(* IEC 61131-3 sources: CS_4_Aufzugsteuerung/src/Stations/CP112/Steuerung/Class/BusInterfaceVARAN (part 2) *)

END_FUNCTION

FUNCTION VIRTUAL GLOBAL BusInterfaceVARAN::UpdateDO
	VAR_INPUT
		pCmd 	            : ^CmdStruct;
		presult 	        : ^results;
	END_VAR
  VAR
    pUPDATEDOCfg      : ^t_UpdateDOCfg;
    pCurrentDO        : ^t_DOCfg;
    changed           : BOOL;

    p_DOSettingsRd    : ^t_VaranDOSettingsRd;
    p_DOSettingsWr    : ^t_VaranDOSettingsWr;
    p_DOSettingsRdWr  : ^t_VaranDOSettingsRdWr;
  END_VAR

  changed := false;
  pUPDATEDOCfg := ((pCmd^.aPara[0])$^t_UpdateDOCfg);

  pResult^.uiLng := 4;

  if CheckHandle(Handle:= pUPDATEDOCfg^.Handle) then

    pCurrentDO := (pUPDATEDOCfg^.Handle)$^t_DOCfg;

    // Check if parameters were changed
    // Read Object
    if pCurrentDO^.RDWR = _BUS_IF_READ then

      if pCurrentDO^.lengthRead <> pUPDATEDOCfg^.ud_length_read  then
        // Check that new DO length is smaller then max DO length
        if pCurrentDO^.maxLengthRead >= pUPDATEDOCfg^.ud_length_read  then
          pCurrentDO^.lengthRead := pUPDATEDOCfg^.ud_length_read;
          changed := true;
        else
          pResult^.aData[0]$t_BusIFRetvalErrorcode := _BUS_IF_RETVAL_ERROR_UPDATEDO_DOLENGTH;
          return;
        end_if;
      end_if;

      if pCurrentDO^.AddrOffsetRead <>  pUPDATEDOCfg^.ud_addressoff_read then
        pCurrentDO^.AddrOffsetRead := pUPDATEDOCfg^.ud_addressoff_read;
        changed := true;
      end_if;

    // Write Object
    elsif pCurrentDO^.RDWR = _BUS_IF_WRITE then

      if pCurrentDO^.lengthWrite <> pUPDATEDOCfg^.ud_length_write  then
        // Check that new DO length is smaller then max DO length
        if pCurrentDO^.maxLengthWrite >= pUPDATEDOCfg^.ud_length_write  then
          pCurrentDO^.lengthWrite := pUPDATEDOCfg^.ud_length_write;
          changed := true;
        else
          pResult^.aData[0]$t_BusIFRetvalErrorcode := _BUS_IF_RETVAL_ERROR_UPDATEDO_DOLENGTH;
          return;
        end_if;
      end_if;

      if pCurrentDO^.AddrOffsetWrite <>  pUPDATEDOCfg^.ud_addressoff_write then
        pCurrentDO^.AddrOffsetWrite := pUPDATEDOCfg^.ud_addressoff_write;
        changed := true;
      end_if;

    // Read Write Object
    else

      if pCurrentDO^.lengthRead <> pUPDATEDOCfg^.ud_length_read  then
        // Check that new DO length is smaller then max DO length
        if pCurrentDO^.maxLengthRead >= pUPDATEDOCfg^.ud_length_read  then
          pCurrentDO^.lengthRead := pUPDATEDOCfg^.ud_length_read;
          changed := true;
        else
          pResult^.aData[0]$t_BusIFRetvalErrorcode := _BUS_IF_RETVAL_ERROR_UPDATEDO_DOLENGTH;
          return;
        end_if;
      end_if;

      if pCurrentDO^.AddrOffsetRead <>  pUPDATEDOCfg^.ud_addressoff_read then
        pCurrentDO^.AddrOffsetRead := pUPDATEDOCfg^.ud_addressoff_read;
        changed := true;
      end_if;

      if pCurrentDO^.lengthWrite <> pUPDATEDOCfg^.ud_length_write  then
        // Check that new DO length is smaller then max DO length
        if pCurrentDO^.maxLengthWrite >= pUPDATEDOCfg^.ud_length_write  then
          pCurrentDO^.lengthWrite := pUPDATEDOCfg^.ud_length_write;
          changed := true;
        else
          pResult^.aData[0]$t_BusIFRetvalErrorcode := _BUS_IF_RETVAL_ERROR_UPDATEDO_DOLENGTH;
          return;
        end_if;
      end_if;

      if pCurrentDO^.AddrOffsetWrite <>  pUPDATEDOCfg^.ud_addressoff_write then
        pCurrentDO^.AddrOffsetWrite := pUPDATEDOCfg^.ud_addressoff_write;
        changed := true;
      end_if;

    end_if;

    if b_PayloadSupport then
      if changed then
        // Update Address and length
        // Read Object
        if pCurrentDO^.RDWR = _BUS_IF_READ then

          ChangeDOLengthOffset( ud_DOHandle     := pCurrentDO^.pHandle$UDINT
                              , ud_offset_read  := pCurrentDO^.AddrOffsetRead
                              , ud_length_read  := pCurrentDO^.lengthRead);

        // Write Object
        elsif pCurrentDO^.RDWR = _BUS_IF_WRITE then

          ChangeDOLengthOffset( ud_DOHandle     := pCurrentDO^.pHandle$UDINT
                              , ud_offset_write := pCurrentDO^.AddrOffsetWrite
                              , ud_length_write := pCurrentDO^.lengthWrite);

        // Read Write Object
        else
          ChangeDOLengthOffset( ud_DOHandle     := pCurrentDO^.pHandle$UDINT
                              , ud_offset_read  := pCurrentDO^.AddrOffsetRead
                              , ud_length_read  := pCurrentDO^.lengthRead
                              , ud_offset_write := pCurrentDO^.AddrOffsetWrite
                              , ud_length_write := pCurrentDO^.lengthWrite);
        end_if;
      end_if;
    elsif pCurrentDO^.IsLongDO = FALSE then

      // Update Address and length and Reset DO
      // Read Object
      if pCurrentDO^.RDWR = _BUS_IF_READ then

        p_DOSettingsRd    := pCurrentDO^.pDataRead$^t_VaranDOSettingsRd  - VM_DO_OFFSET_RD;

        p_DOSettingsRd^.ud_Address                := DeviceAddress + pCurrentDO^.AddrOffsetRead;
        p_DOSettingsRd^.us_ByteCnt                := pCurrentDO^.lengthRead$USINT;
        pCurrentDO^.pHandle^.usLengthofExpAnswer  := sizeof(t_VaranDOSettingsRd.us_Command) + pCurrentDO^.lengthRead;

        ResetDataObject(p_handleDO:=  pCurrentDO^.pHandle
                      , us_state  :=  pCurrentDO^.pHandle^.ucCtrlStat AND 3         // don't change run status, just recalculate the retry timeout here
                      , ud_bytes  :=  pCurrentDO^.lengthRead);

      // Write Object
      elsif pCurrentDO^.RDWR = _BUS_IF_WRITE then

        p_DOSettingsWr    := pCurrentDO^.pDataWrite$^t_VaranDOSettingsWr - VM_DO_OFFSET_WR;

        p_DOSettingsWr^.ud_Address              := DeviceAddress + pCurrentDO^.AddrOffsetWrite;
        p_DOSettingsWr^.us_ByteCnt              := pCurrentDO^.lengthWrite$USINT;
        pCurrentDO^.pHandle^.usSendBufferLength := sizeof(t_VaranDOSettingsWr) + pCurrentDO^.lengthWrite;

        ResetDataObject(p_handleDO:=  pCurrentDO^.pHandle
                      , us_state  :=  pCurrentDO^.pHandle^.ucCtrlStat AND 3         // don't change run status, just recalculate the retry timeout here
                      , ud_bytes  :=  pCurrentDO^.lengthWrite);

      // Read Write Object
      else
        p_DOSettingsRdWr  := pCurrentDO^.pDataWrite$^t_VaranDOSettingsRdWr - VM_DO_OFFSET_RDWR;

        p_DOSettingsRdWr^.ud_AddressRd := DeviceAddress + pCurrentDO^.AddrOffsetRead;
        p_DOSettingsRdWr^.ud_AddressWr := DeviceAddress + pCurrentDO^.AddrOffsetWrite;

        p_DOSettingsRdWr^.us_ByteCntRd  := pCurrentDO^.lengthRead$USINT;
        p_DOSettingsRdWr^.us_ByteCntWr  := pCurrentDO^.lengthWrite$USINT;

        pCurrentDO^.pHandle^.usLengthofExpAnswer  := sizeof(t_VaranDOSettingsRdWr.us_Command) + pCurrentDO^.lengthRead;
        pCurrentDO^.pHandle^.usSendBufferLength   := sizeof(t_VaranDOSettingsRdWr) + pCurrentDO^.lengthWrite;

        ResetDataObject(p_handleDO:=  pCurrentDO^.pHandle
                      , us_state  :=  pCurrentDO^.pHandle^.ucCtrlStat AND 3         // don't change run status, just recalculate the retry timeout here
                      , ud_bytes  :=  pCurrentDO^.lengthRead + pCurrentDO^.lengthWrite);

      end_if;
    else

      // change long DO

      // Update Address and length and Reset DO
      // Read Object
      if pCurrentDO^.RDWR = _BUS_IF_READ then

        pCurrentDO^.pLongDOSettings^.ud_Address      := DeviceAddress + pCurrentDO^.AddrOffsetRead;
        pCurrentDO^.pLongDOSettings^.ui_ByteCount0   := pCurrentDO^.lengthRead;
        pCurrentDO^.pLongDOSettings^.us_ByteCount1   := 0;
        pCurrentDO^.pHandle^.usSendBufferLength      := 16#FFFF;
        pCurrentDO^.pHandle^.usLengthofExpAnswer     := 16#FFFF;

      // Write Object
      elsif pCurrentDO^.RDWR = _BUS_IF_WRITE then

        pCurrentDO^.pLongDOSettings^.ud_Address      := DeviceAddress + pCurrentDO^.AddrOffsetWrite;
        pCurrentDO^.pLongDOSettings^.ui_ByteCount0   := pCurrentDO^.lengthWrite;
        pCurrentDO^.pLongDOSettings^.us_ByteCount1   := 0;
        pCurrentDO^.pHandle^.usSendBufferLength      := 16#FFFF;
        pCurrentDO^.pHandle^.usLengthofExpAnswer     := 16#FFFF;

      end_if;
    end_if;

    pResult^.aData[0]$t_BusIFRetvalErrorcode := _BUS_IF_RETVAL_OK;

  else
    pResult^.aData[0]$t_BusIFRetvalErrorcode := _BUS_IF_RETVAL_ERROR_INVALID_HANDLE;
  end_if;

END_FUNCTION

FUNCTION VIRTUAL GLOBAL BusInterfaceVARAN::UpdateMoveDO
	VAR_INPUT
		pCmd 	        : ^CmdStruct;
		presult 	    : ^results;
	END_VAR
  VAR
    pUPDATEDOCfg  : ^t_UpdateDOMoveCfg;
    pCurrentDO    : ^t_DOMoveCfg;
    sd_retval     : DINT;
  END_VAR

  pUPDATEDOCfg := ((pCmd^.aPara[0])$^t_UpdateDOMoveCfg);

  pResult^.uiLng := 4;

  if CheckMovHandle(Handle:= pUPDATEDOCfg^.Handle) then

    pCurrentDO := (pUPDATEDOCfg^.Handle)$^t_DOMoveCfg;

    // Check if length Parameter was passed
    // Length is used with Payload and without
    if (pUPDATEDOCfg^.ud_length_move <> 0) &
       pUPDATEDOCfg^.ud_length_move <> VM_DO_PROPERTY_INVALID  then
      // if the size is smaller than the maximum or if we don't have interrupted our own copy for the move command
      if (pUPDATEDOCfg^.ud_length_move <= pCurrentDO^.lengthMoveMax) | (us_SkippedWriteBlocks = 0) then
        pCurrentDO^.lengthMove := pUPDATEDOCfg^.ud_length_move;
      else
        pResult^.aData[0]$t_BusIFRetvalErrorcode := _BUS_IF_RETVAL_ERROR_UPDATEDO_DOLENGTH;
        return;
      end_if;
    end_if;

    if b_PayloadSupport then

      if  pUPDATEDOCfg^.ud_handle_source <> 0 &
          pUPDATEDOCfg^.ud_handle_source <> VM_DO_PROPERTY_INVALID  then

        pCurrentDO^.sourceDOHandle := pUPDATEDOCfg^.ud_handle_source;
      end_if;

      if  pUPDATEDOCfg^.ud_addressoff_source <> VM_DO_PROPERTY_INVALID  then  // 0 is valid offset

        pCurrentDO^.sourceDOOffset := pUPDATEDOCfg^.ud_addressoff_source;
      end_if;

      if  pUPDATEDOCfg^.ud_handle_dest <> 0 &
          pUPDATEDOCfg^.ud_handle_dest <> VM_DO_PROPERTY_INVALID  then

        pCurrentDO^.destDOHandle := pUPDATEDOCfg^.ud_handle_dest;
      end_if;

      if  pUPDATEDOCfg^.ud_addressoff_dest <> VM_DO_PROPERTY_INVALID  then  // 0 is valid offset

        pCurrentDO^.destDOOffset := pUPDATEDOCfg^.ud_addressoff_dest;
      end_if;

      sd_retval := ChangeMovDOLengthOffset( ud_MovDOHandle              := pCurrentDO^.pHandle$UDINT
                                          , ud_SourceReadDOHandle       := pCurrentDO^.sourceDOHandle
                                          , ud_SourceReadOffset         := pCurrentDO^.sourceDOOffset
                                          , ud_DestinationWriteDOHandle := pCurrentDO^.destDOHandle
                                          , ud_DestinationWriteOffset   := pCurrentDO^.destDOOffset
                                          , ud_LengthMove               := pCurrentDO^.lengthMove);

      if sd_retval then
        pResult^.aData[0]$t_BusIFRetvalErrorcode := _BUS_IF_RETVAL_ERROR_UPDATE_MOVE_DO_FAILED;
      else
        pResult^.aData[0]$t_BusIFRetvalErrorcode := _BUS_IF_RETVAL_OK;
      end_if;

    else

      if pUPDATEDOCfg^.p_sourcedata <> nil &
         pUPDATEDOCfg^.p_sourcedata <> VM_DO_PROPERTY_INVALID then

        pCurrentDO^.pSourceDOData := pUPDATEDOCfg^.p_sourcedata;
      end_if;

      if pUPDATEDOCfg^.p_destdata   <> nil &
         pUPDATEDOCfg^.p_destdata   <> VM_DO_PROPERTY_INVALID then

        pCurrentDO^.pDestDOData := pUPDATEDOCfg^.p_destdata;
      end_if;

      pCurrentDO^.p_MovSettings^.ud_AddressSrc  := pCurrentDO^.pSourceDOData$UDINT;
      pCurrentDO^.p_MovSettings^.ud_AddressDest := pCurrentDO^.pDestDOData$UDINT;
      pCurrentDO^.p_MovSettings^.ui_ByteCnt     := pCurrentDO^.lengthMove;

      pResult^.aData[0]$t_BusIFRetvalErrorcode := _BUS_IF_RETVAL_OK;
    end_if;

  else
    pResult^.aData[0]$t_BusIFRetvalErrorcode := _BUS_IF_RETVAL_ERROR_INVALID_HANDLE;
  end_if;

END_FUNCTION

FUNCTION VIRTUAL GLOBAL BusInterfaceVARAN::SetDOPrescaler
	VAR_INPUT
		pCmd 	        : ^CmdStruct;
		presult 	    : ^results;
	END_VAR
  VAR
    pSetDOPreSCfg : ^t_SetDoPrescaler;
    pCurrentDO    : ^t_DOCfg;
  END_VAR

  pSetDOPreSCfg := ((pCmd^.aPara[0])$^t_SetDoPrescaler);

  pResult^.uiLng := 4;

  if CheckHandle(Handle:= pSetDOPreSCfg^.Handle) then

    pCurrentDO := (pSetDOPreSCfg^.Handle)$^t_DOCfg;

    if b_PayloadSupport then

      if SetPrescaler( ud_DOHandle   := pCurrentDO^.pHandle$UDINT
                     , Prescaler     := pSetDOPreSCfg^.Prescaler
                     , PrescalerCnt  := 0) = VARANMANAGER_OK then // Start at 0 = default We probably need to extend this functionality

        pResult^.aData[0]$t_BusIFRetvalErrorcode := _BUS_IF_RETVAL_OK;
      else
        pResult^.aData[0]$t_BusIFRetvalErrorcode := _BUS_IF_RETVAL_ERROR_INVALID_HANDLE;
      end_if;
    else

      pCurrentDO^.pHandle^.ucExePrescaler := pSetDOPreSCfg^.Prescaler;
      pCurrentDO^.PreScaler := pSetDOPreSCfg^.Prescaler;  // Saved as needed again as init value

      pResult^.aData[0]$t_BusIFRetvalErrorcode := _BUS_IF_RETVAL_OK;
    end_if;
  else

    pResult^.aData[0]$t_BusIFRetvalErrorcode := _BUS_IF_RETVAL_ERROR_INVALID_HANDLE;
  end_if;

END_FUNCTION

FUNCTION VIRTUAL GLOBAL BusInterfaceVARAN::SetTasksPrescaler
	VAR_INPUT
		pCmd 	            : ^CmdStruct;
		presult 	        : ^results;
	END_VAR
  VAR
  	pTaskPreScalerCfg : ^t_TaskPreScaler;
  END_VAR

  pTaskPreScalerCfg  := ((pCmd^.aPara[0])$^t_TaskPreScaler);

  pResult^.uiLng := 4;

  // Check passed data
  if pTaskPreScalerCfg^.Prescaler > 0 &
     pTaskPreScalerCfg^.Prescaler >= pTaskPreScalerCfg^.RtPreScanTrigger &
     pTaskPreScalerCfg^.Prescaler >= pTaskPreScalerCfg^.RtPostScanTrigger &
     pTaskPreScalerCfg^.Prescaler >= pTaskPreScalerCfg^.CyTrigger then

    TaskPrescaler.MaxCnt            := pTaskPreScalerCfg^.Prescaler;
    TaskPrescaler.RtPreScanTigger   := pTaskPreScalerCfg^.RtPreScanTrigger;
    TaskPrescaler.RtPostScanTrigger := pTaskPreScalerCfg^.RtPostScanTrigger;
    TaskPrescaler.CyTrigger         := pTaskPreScalerCfg^.CyTrigger;

    pResult^.aData[0]$t_BusIFRetvalErrorcode := _BUS_IF_RETVAL_OK;
  else
    pResult^.aData[0]$t_BusIFRetvalErrorcode := _BUS_IF_RETVAL_ERROR_INVALID_DATA;
  end_if;

END_FUNCTION

FUNCTION VIRTUAL GLOBAL BusInterfaceVARAN::ResetDO
	VAR_INPUT
		pCmd 	      : ^CmdStruct;
		presult 	  : ^results;
	END_VAR
  VAR
    pResetDOCfg : ^t_ResetDOCfg;
    pCurrentDO  : ^t_DOCfg;
  END_VAR

  pResult^.uiLng := 4;

  pResetDOCfg := ((pCmd^.aPara[0])$^t_ResetDOCfg);

  if CheckHandle(Handle:= pResetDOCfg^.Handle) then

    // Paylaod DO auto calculate Timeout when the DO changes
    // Just return OK
    if b_PayloadSupport = false then

      pCurrentDO := (pResetDOCfg^.Handle)$^t_DOCfg;

      // Reset DO
      // Read Object
      if (pCurrentDO^.RDWR = _BUS_IF_READ) then
        if pCurrentDO^.IsLongDO then
          ResetDataObject(p_handleDO :=  pCurrentDO^.pHandle
                          , us_state :=  VARAN_DO_NO_RUN         // No auto run, DO must be started by specific command
                          , ud_bytes :=  128);
        else
          ResetDataObject(p_handleDO :=  pCurrentDO^.pHandle
                          , us_state :=  VARAN_DO_NO_RUN         // No auto run, DO must be started by specific command
                          , ud_bytes :=  pCurrentDO^.lengthRead);
        end_if;

      // Write DO
      elsif pCurrentDO^.RDWR = _BUS_IF_WRITE then
        if pCurrentDO^.IsLongDO then
          ResetDataObject(p_handleDO :=  pCurrentDO^.pHandle
                          , us_state :=  VARAN_DO_NO_RUN         // No auto run, DO must be started by specific command
                          , ud_bytes :=  128);
        else
          ResetDataObject(p_handleDO :=  pCurrentDO^.pHandle
                          , us_state :=  VARAN_DO_NO_RUN         // No auto run, DO must be started by specific command
                          , ud_bytes :=  pCurrentDO^.lengthWrite);
        end_if;

      // Read Write DO
      else

        ResetDataObject(p_handleDO:=  pCurrentDO^.pHandle
                        , us_state  :=  VARAN_DO_NO_RUN         // No auto run, DO must be started by specific command
                        , ud_bytes  :=  pCurrentDO^.lengthRead + pCurrentDO^.lengthWrite);

      end_if;

    end_if;

    pResult^.aData[0]$t_BusIFRetvalErrorcode := _BUS_IF_RETVAL_OK;

  else
    pResult^.aData[0]$t_BusIFRetvalErrorcode := _BUS_IF_RETVAL_ERROR_INVALID_HANDLE;
  end_if;

END_FUNCTION

FUNCTION VIRTUAL GLOBAL BusInterfaceVARAN::AddTask
	VAR_INPUT
		pCmd 	        : ^CmdStruct;
		presult       : ^results;
	END_VAR
  VAR
  	pTASKCfg      : ^t_TaskCfg;
    _ud_dol_type  : UDINT;
  END_VAR

  presult^.uiLng    := 4;

  pTASKCfg := ((pCmd^.aPara[0])$^t_TaskCfg);

  // Check for null pointer
  if pTASKCfg^.pthis then

        // Convert passed t_BusIFPriority  to VARAN ud_dol_type
    if pTASKCfg^.Priority = _BUS_IF_ISO then
      _ud_dol_type := VARAN_DOL_ISO;
    else
      _ud_dol_type := VARAN_DOL_ASY;
    end_if;

    // Save the passed callback pointer according to the callOptions
    if pTASKCfg^.callOptions = CALL_OPTION_RT_PRESCAN then
      p_UserCalls.p_UpdateRt := (pTASKCfg^.pthis)$pVirtualBase;
    elsif pTASKCfg^.callOptions = CALL_OPTION_RT_POSTSCAN then
      p_UserCalls.p_UpDateRtPostScan := (pTASKCfg^.pthis)$pVirtualBase;
    elsif pTASKCfg^.callOptions = (CALL_OPTION_RT_PRESCAN or CALL_OPTION_RT_POSTSCAN) then
      p_UserCalls.p_UpdateRt := (pTASKCfg^.pthis)$pVirtualBase;
      p_UserCalls.p_UpDateRtPostScan := (pTASKCfg^.pthis)$pVirtualBase;
    else
      p_UserCalls.p_UpdateCy := (pTASKCfg^.pthis)$pVirtualBase;
    end_if;

    //Install Varantask
    VaranIn.AddVaranTask( _ud_dol_type,
                          p_this:=this,       // The callback pointer cannot be used directly because the class must be derived from VaranBase (p_VaranBase)
                          pTASKCfg^.callOptions);

    pResult^.aData[0]$t_BusIFRetvalErrorcode := _BUS_IF_RETVAL_OK;
  else
    pResult^.aData[0]$t_BusIFRetvalErrorcode := _BUS_IF_RETVAL_ERROR_INVALID_POINTER;
  end_if;

END_FUNCTION

FUNCTION VIRTUAL GLOBAL BusInterfaceVARAN::SetRunState
	VAR_INPUT
		pCmd 	            : ^CmdStruct;
		presult 	        : ^results;
	END_VAR
  VAR
  	pSETRUNSTATECfg   : ^t_SetRunStateCfg;
    pCurrentDO        : ^t_DOCfg;
    pCurrentDOMove    : ^t_DOMoveCfg;
    sd_RetVal         : DINT;
  END_VAR

  presult^.uiLng  := 4;

  pSETRUNSTATECfg := ((pCmd^.aPara[0])$^t_SetRunStateCfg);

  // Standard DO -----------------------------------------------------------------------------
  if CheckHandle(Handle:= pSETRUNSTATECfg^.Handle) then

    pCurrentDO := (pSETRUNSTATECfg^.Handle)$^t_DOCfg;

    if b_PayloadSupport then
      if pSETRUNSTATECfg^.NewRunState = _BUS_IF_RUN_STATE_SINGLE_RUN then
        pCurrentDO^.b_DOIsRunning.ContRun       := false; // Override cont run
        pCurrentDO^.b_DOIsRunning.StartRequest  := true;
        pResult^.aData[0]$t_BusIFRetvalErrorcode := _BUS_IF_RETVAL_OK;
      elsif pSETRUNSTATECfg^.NewRunState = _BUS_IF_RUN_STATE_CONT_RUN then
        if EnableDO(ud_DOHandle := pCurrentDO^.pHandle$UDINT) = VARANMANAGER_OK then

          //check if do must be added to list
          if bAddDOsToListSupport
          & pCurrentDO^.bsDoInsert.DOisInserted = FALSE
          & pCurrentDO^.bsDoInsert.RequestInsertLater = TRUE then
            sd_RetVal := MULTI_VARAN_IINSERTDOINTODOL(pCurrentDO^.pHandle$UDINT);
            pCurrentDO^.bsDoInsert.DOisInserted := TRUE;
          end_if;

          pResult^.aData[0]$t_BusIFRetvalErrorcode := _BUS_IF_RETVAL_OK;
        else
          pResult^.aData[0]$t_BusIFRetvalErrorcode := _BUS_IF_RETVAL_ERROR_INVALID_HANDLE;
        end_if;
        pCurrentDO^.b_DOIsRunning         := 0; // Override any singlerun states
        pCurrentDO^.b_DOIsRunning.ContRun := true;
      else
        if DisableDO(ud_DOHandle := pCurrentDO^.pHandle$UDINT) = VARANMANAGER_OK then
          pResult^.aData[0]$t_BusIFRetvalErrorcode := _BUS_IF_RETVAL_OK;
        else
          pResult^.aData[0]$t_BusIFRetvalErrorcode := _BUS_IF_RETVAL_ERROR_INVALID_HANDLE;
        end_if;
        pCurrentDO^.b_DOIsRunning         := 0;
      end_if;
    else
      if pSETRUNSTATECfg^.NewRunState = _BUS_IF_RUN_STATE_SINGLE_RUN then
        pCurrentDO^.pHandle^.ucCtrlStat := SetRunStatus(state:=VARAN_DO_SINGLE_RUN);
      elsif pSETRUNSTATECfg^.NewRunState = _BUS_IF_RUN_STATE_CONT_RUN then
        pCurrentDO^.pHandle^.ucCtrlStat := SetRunStatus(state:=VARAN_DO_CONT_RUN);
      else
        pCurrentDO^.pHandle^.ucCtrlStat := SetRunStatus(state:=VARAN_DO_NO_RUN);
      end_if;

      pResult^.aData[0]$t_BusIFRetvalErrorcode := _BUS_IF_RETVAL_OK;
    end_if;

  // Move DO ----------------------------------------------------------------------------------------
  elsif CheckMovHandle(Handle:= pSETRUNSTATECfg^.Handle) then

    pCurrentDOMove := (pSETRUNSTATECfg^.Handle)$^t_DOMoveCfg;

    if b_PayloadSupport then
      if pSETRUNSTATECfg^.NewRunState = _BUS_IF_RUN_STATE_SINGLE_RUN then
        pCurrentDOMove^.b_DOIsRunning.ContRun       := false; // Override cont run
        pCurrentDOMove^.b_DOIsRunning.StartRequest  := true;
        pResult^.aData[0]$t_BusIFRetvalErrorcode := _BUS_IF_RETVAL_OK;
      elsif pSETRUNSTATECfg^.NewRunState = _BUS_IF_RUN_STATE_CONT_RUN then
        if EnableDO(ud_DOHandle := pCurrentDOMove^.pHandle$UDINT) = VARANMANAGER_OK then
          pResult^.aData[0]$t_BusIFRetvalErrorcode := _BUS_IF_RETVAL_OK;
        else
          pResult^.aData[0]$t_BusIFRetvalErrorcode := _BUS_IF_RETVAL_ERROR_INVALID_HANDLE;
        end_if;
        pCurrentDOMove^.b_DOIsRunning         := 0; // Override any singlerun states
        pCurrentDOMove^.b_DOIsRunning.ContRun := true;
      else
        if DisableDO(ud_DOHandle := pCurrentDOMove^.pHandle$UDINT) = VARANMANAGER_OK then
          pResult^.aData[0]$t_BusIFRetvalErrorcode := _BUS_IF_RETVAL_OK;
        else
          pResult^.aData[0]$t_BusIFRetvalErrorcode := _BUS_IF_RETVAL_ERROR_INVALID_HANDLE;
        end_if;
        pCurrentDOMove^.b_DOIsRunning         := 0;
      end_if;
    else
      if pSETRUNSTATECfg^.NewRunState = _BUS_IF_RUN_STATE_SINGLE_RUN then
        pCurrentDOMove^.pHandle^.ucCtrlStat := SetRunStatus(state:=VARAN_DO_SINGLE_RUN);
      elsif pSETRUNSTATECfg^.NewRunState = _BUS_IF_RUN_STATE_CONT_RUN then
        pCurrentDOMove^.pHandle^.ucCtrlStat := SetRunStatus(state:=VARAN_DO_CONT_RUN);
      else
        pCurrentDOMove^.pHandle^.ucCtrlStat := SetRunStatus(state:=VARAN_DO_NO_RUN);
      end_if;

      pResult^.aData[0]$t_BusIFRetvalErrorcode := _BUS_IF_RETVAL_OK;
    end_if;

  else
    pResult^.aData[0]$t_BusIFRetvalErrorcode := _BUS_IF_RETVAL_ERROR_INVALID_HANDLE;
  end_if;

END_FUNCTION

FUNCTION VIRTUAL GLOBAL BusInterfaceVARAN::SetSyncData
	VAR_INPUT
		pCmd 	        : ^CmdStruct;
		presult 	    : ^results;
	END_VAR
  VAR
    pSYNCDATACfg  :  ^t_SyncData;
    i             : USINT;
  END_VAR

  presult^.uiLng  := 4;

  pSYNCDATACfg    := ((pCmd^.aPara[0])$^t_SyncData);

  i := pSYNCDATACfg^.us_sync_nr;

  if  i >= 0 &
      i <  4 then

    SyncData[i].us_sync_nr                := pSYNCDATACfg^.us_sync_nr;
    SyncData[i].sd_offset                 := pSYNCDATACfg^.sd_offset;
    SyncData[i].us_period_multiplier      := pSYNCDATACfg^.us_period_multiplier;
    SyncData[i].us_enable_frame_count     := pSYNCDATACfg^.us_enable_frame_count;
    SyncData[i].us_frame_count_threshold  := pSYNCDATACfg^.us_frame_count_threshold;
    SyncData[i].b_use_divider_sync        := pSYNCDATACfg^.b_use_divider_sync;

    bSetPll := TRUE;

    pResult^.aData[0]$t_BusIFRetvalErrorcode := _BUS_IF_RETVAL_OK;
  else
    pResult^.aData[0]$t_BusIFRetvalErrorcode := _BUS_IF_RETVAL_ERROR_INVALID_SYNC;
  end_if;

END_FUNCTION

FUNCTION VIRTUAL BusInterfaceVARAN::CheckHandle
	VAR_INPUT
		Handle 	    : UDINT;
	END_VAR
	VAR_OUTPUT
		IsOk 	      : BOOL;
	END_VAR
  VAR
    ListOffset  : UDINT;
  END_VAR

  IsOk := false;

  // Handle must be not nil and there must be elements in the array.
  if Handle & NrDO then
    ListOffset := (Handle - (#DOList[0])$UDINT);
    if ((ListOffset MOD sizeof(t_DOCfg)) = 0) & ((ListOffset/sizeof(t_DOCfg)) < NrDO) then
      IsOk := true;
    end_if;
  end_if;

END_FUNCTION

FUNCTION VIRTUAL BusInterfaceVARAN::CheckMovHandle
	VAR_INPUT
		Handle 	    : UDINT;
	END_VAR
	VAR_OUTPUT
		IsOk 	      : BOOL;
	END_VAR
  VAR
    ListOffset  : UDINT;
  END_VAR

  IsOk := false;

  // Handle must be not nil and there must be elements in the array.
  if Handle & NrDOMove then
    ListOffset := (Handle - (#DOListMove[0])$UDINT);
    if ((ListOffset MOD sizeof(t_DOMoveCfg)) = 0) & ((ListOffset/sizeof(t_DOMoveCfg)) < NrDOMove) then
      IsOk := true;
    end_if;
  end_if;

END_FUNCTION

FUNCTION VIRTUAL GLOBAL BusInterfaceVARAN::UpdateRetryCounter
  VAR
    i                 : USINT;
	  tempRetryCounter  : USINT;
    pDOElement        : ^t_DOCfg;
  END_VAR

  // Standard DOs --------------------------------------------------------------------------
  if NrDO then
    pDOElement := #DOList[0];
    for i := 0 to (NrDO - 1) do

      tempRetryCounter := GetRetryCounter(ud_DOHandle := pDOElement^.pHandle$UDINT);

      if ( tempRetryCounter <> pDOElement^.OldRetryCounter) then
        RetryCounter += TO_USINT( tempRetryCounter - pDOElement^.OldRetryCounter );
        pDOElement^.OldRetryCounter := tempRetryCounter;
      end_if;

      pDOElement += sizeof(t_DOCfg);
    end_for;
  end_if;

END_FUNCTION

FUNCTION BusInterfaceVARAN::BusInterfaceVARAN
	VAR_OUTPUT
		ret_code 	: ConfStates;
	END_VAR

  ui_PostInitIndex := 16#FFFF;

  // initialize with 0xff for invalid
  _memset(dest:=#SyncData, usByte:=16#FF, cntr:=sizeof(SyncData));

  if OS_CILGet(INTERFACE_VARANMANAGER, #pVaran) <> SYS_ERR_NONE then
    LogError("@0196 (BusInterfaceVARAN::BusInterfaceVARAN) Failed to get VARAN-CIL (interface to OS)!");
  end_if;

  b_LongDOsPossible := GetLongDOsPossible();

	ret_code := C_OK;

END_FUNCTION

FUNCTION VIRTUAL GLOBAL BusInterfaceVARAN::Varan_HwInterrupt
	VAR_INPUT
		ud_reason 	: UDINT;
		ud_data 	  : ^t_CallBackInterrupt;
	END_VAR
	VAR_OUTPUT
		sd_retval 	: DINT;
	END_VAR
  VAR
  	tempCmd     : CmdStruct;
    _result     : results;
  END_VAR;

  // Turn off DO's
  SetDOsOff();

  // Check for 0 pointer
  if p_UserCalls.p_Callback then
    // Call the corrosponding function in the operator class
    tempCmd.uiCmd := _BUS_IF_HWINTERRUPT;
    p_UserCalls.p_Callback^.pSvrChCmd.NewInst(#tempCmd,#_result);
  end_if;
  sd_retval := Varan_Base::Varan_HwInterrupt(ud_reason, ud_data);

END_FUNCTION

FUNCTION VIRTUAL BusInterfaceVARAN::LogErrorExt
	VAR_INPUT
		e_msg 	    : ^CHAR;
		p_extThis1 	: pVirtualBase;
		p_extThis2 	: pVirtualBase;
	END_VAR
  VAR
    sz_name     : ARRAY [ 0..255 ] OF CHAR;
    MyMsg       : ARRAY [0..599] OF CHAR;
  END_VAR

  if p_extThis1 = nil then
    p_extThis1 := this;
  end_if;

  if p_extThis2 then
    _GetObjName( p_extThis2, #sz_name[ 0 ] );
#ifdef HWC_LimitObjName
    HWC_LimitObjName(#sz_name[ 0 ]);
#endif
    _strncpy(dest:=#MyMsg[0], src:=e_msg, max:=200);
    _strcat( dest:=#MyMsg[0], src:=" ");
    _strcat( dest:=#MyMsg[0], src:=#sz_name[0]);

#ifdef HWC_LogError
    HWC_LogError(p_extThis1, #MyMsg[0]);
#endif

  else
#ifdef HWC_LogError
    HWC_LogError(p_extThis1, e_msg);
#endif
  end_if;

END_FUNCTION

FUNCTION VIRTUAL BusInterfaceVARAN::InstallCallbackObject
	VAR_OUTPUT
		sd_retval 	: DINT;
	END_VAR

  // we don't install the callback here (1st init). it's installed in the 2nd init, because in the first init the operator may set us to required
  sd_retval := VARANMANAGER_OK;

END_FUNCTION

FUNCTION VIRTUAL BusInterfaceVARAN::GetLongDOsPossible
	VAR_OUTPUT
		LongDOsPossible 	  : BOOL;
	END_VAR
  VAR
    pSPCIInfo           : ^LSL_SPCIINFO;
  	p_sigmatek_devinfo 	: ^PCICONFDATA;
    p_NodeInfo          : ^LSL_VARANNODEINFO;
    ManagerNodeString   : USINT;
    ud_VMNodeHandle     : UDINT;
    s_NodeInfo          : LSL_VARANNODEINFO;
    sd_retval           : DINT;
  END_VAR

  LongDOsPossible := FALSE;

  // check if long DOs are supported by VARAN Manager. Version of wb_varan_manager_control_status_info (Device Type x"0212" of info block) has to be >= 16#25.
  if OS_CILGET( "PCICONFIG", #pSPCIInfo ) =  SYS_ERR_NONE then
    p_sigmatek_devinfo 	:= SPCIINFO_FINDDEVICE(0x0212, 0);
    if p_sigmatek_devinfo = NIL then
      p_sigmatek_devinfo 	:= SPCIINFO_FINDDEVICE(0x0214, 0); //check for new varan interface
    end_if;
    // check if the Manager supports LongDOs
    if p_sigmatek_devinfo & (p_sigmatek_devinfo^.Version >= 16#25) then
      LongDOsPossible := TRUE;
    else
      // we don't get the device at a c-ipc, because it's a pci plug-in card
      if pVaran & (_WhoAmI = DESTPLC_C_IPC) then
        // now check the platform and the corresponding fpga version

        //get manager node info from os
        ManagerNodeString := 0;

        //call OS - function (must be OS-funciton because of error handling)
        if b_PayloadSupport then
          // Get the Handle of the VM
          sd_retval := MULTI_VARAN_iGetNodeHandle(udManagerNumber := ud_VaranManagerNr
                                                , pszHardwarePath := #ManagerNodeString
                                                , phNodeHandle    := #ud_VMNodeHandle);

          if sd_retval = VARANMANAGER_OK then
            p_NodeInfo := #s_NodeInfo;
            sd_retval := MULTI_VARAN_iGetNodeInformation( hNodeHandle := ud_VMNodeHandle
                                                        , psNodeInfo  := p_NodeInfo);     // Pass a pointer to the buffer into which the data will be written, instead of getting a pointer to te data
          end_if;

        else
          sd_retval := VARAN_iGetNodeInfo(uiManager	:= ud_VaranManagerNr
                                        , pucNode	  := #ManagerNodeString
                                        , pNodeInfo	:= #p_NodeInfo
                                        );
        end_if;

        if	( sd_retval = VARANMANAGER_OK ) & p_NodeInfo then
          case p_NodeInfo^.uiDeviceID of
            1000: // VM051    >= 1.6
              if p_NodeInfo^.ucFPGAVersion >= 16#16 then
                LongDOsPossible := TRUE;
              end_if;

            1030, // VM052    >= 1.4
            1150: // VM052-1  same fpga file
              if p_NodeInfo^.ucFPGAVersion >= 16#14 then
                LongDOsPossible := TRUE;
              end_if;

            1031: // VM052H   not necessary, this card doesn't work on a C-IPC (created for customer specific hardware)

            1044: // VMC052   >= 1.3
              if p_NodeInfo^.ucFPGAVersion >= 16#13 then
                LongDOsPossible := TRUE;
              end_if;

            1063, // VM052-3  >= 1.4
            1093: // VM053    same fpga file
              if p_NodeInfo^.ucFPGAVersion >= 16#14 then
                LongDOsPossible := TRUE;
              end_if;

            1080: // VM052-4  no fpga available

          end_case;
        end_if;
      end_if;
    end_if;
  end_if;

END_FUNCTION

FUNCTION VIRTUAL GLOBAL BusInterfaceVARAN::Varan_HwSubBusReady
	VAR_INPUT
		ud_data 	  : UDINT;
	END_VAR
	VAR_OUTPUT
		sd_retval 	: DINT;
	END_VAR
  VAR
  	tempCmd     : CmdStruct;
    _result     : results;
  END_VAR

  // Check for 0 pointer
  if p_UserCalls.p_Callback then
    // Call the corresponding function in the operator class
    tempCmd.uiCmd := _BUS_IF_HWSUB_BUS_READY;
    p_UserCalls.p_Callback^.pSvrChCmd.NewInst(#tempCmd,#_result);

    sd_retval := _result.aData[0]$DINT;
  else
    sd_retval := 0;
  end_if;

END_FUNCTION

FUNCTION VIRTUAL GLOBAL BusInterfaceVARAN::State::NewInst
	VAR_INPUT
		pPara 	    : ^CmdStruct;
		pResult 	  : ^Results;
	END_VAR
	VAR_OUTPUT
		ret_code 	  : IprStates;
	END_VAR
  VAR
  	tempCmd     : CmdStruct;
    _result     : results;
    // local variables for the Requested HWTString
    pStr_HWTRequested       : ^CHAR;
    us_HWTRequestedCurrIndex: USINT;
    pStr_HWTreenEntry       : ^CHAR;
    ud_HWCRetcode           : t_HWCRetvalReturnCode;
    b_CallThisModule        : BOOL;
  END_VAR

  pStr_HWTRequested         := NIL;
  us_HWTRequestedCurrIndex  := 0;
  pStr_HWTreenEntry         := NIL;
  ud_HWCRetcode             := _HWC_RETVAL_ERROR;
  b_CallThisModule          := TRUE;

	ret_code := READY;

  CASE pPara^.uiCmd OF
//**********************************************************************************************************************************************************
    CMD_POST_INIT_RT_READY:
      // check if operator is ready
      tempCmd.uiCmd := _BUS_IF_POST_INIT_RT_READY;
      ret_code := p_UserCalls.p_Callback^.pSvrChCmd.NewInst(#tempCmd, #_result);

      if bSimulateSDIASManager then

        // if we got an error => return it
        if eSdiasManagerInitSSW = _ErrorOccured then
          ret_code := ERROR;

        //if we're not ready, return busy
        elsif eSdiasManagerInitSSW <> _InitFinished then
          ret_code := BUSY;
        end_if;

      end_if;

//**********************************************************************************************************************************************************
    CMD_GET_HARDWARE_DIAGNOSIS:

      pResult^.aData$t_HWCGetHardwareDiagnosisOut.retcode := _HWC_RETVAL_ERROR_CLASS_NOT_ONLINE;
      ret_code := ERROR;

      pResult^.aData[0]$t_HWCGetHardwareDiagnosisOut.retcode := _HWC_RETVAL_ERROR;

      pStr_HWTRequested := pPara^.aPara[0]$t_HWCGetHardwareDiagnosisIn.pStr_HardewareTreeEntry;

      // Check HWT String
      if pStr_HWTRequested then

        us_HWTRequestedCurrIndex  := pPara^.aPara[0]$t_HWCGetHardwareDiagnosisIn.us_current_index;

        // Check for any Escape sequence
        if (pStr_HWTRequested + us_HWTRequestedCurrIndex)^ and HWT_ESCAPE_SEQU then

          // Check if current index + 1 is valid, pStr_HWTRequested^ + 1 for extra byte of length
          if (us_HWTRequestedCurrIndex + 1) <= (pStr_HWTRequested$^UINT^ + 1) then
            // Update Current index to next position = Place of SDIAS Module
            pPara^.aPara[0]$t_HWCGetHardwareDiagnosisIn.us_current_index   += 1;
            pPara^.aPara[0]$t_HWCGetHardwareDiagnosisIn.us_current_length  -= 1;

            if p_UserCalls.p_Callback then
              ret_code := p_UserCalls.p_Callback^.pSvrChCmd.NewInst(pPara,pResult); //Pass on command to connected extension module
            end_if;

          end_if;

        else
          ret_code := Varan_Base::State.NewInst(pPara, pResult);  // Pass on command to base

          // Call conneceted Class for additional info
          if p_UserCalls.p_Callback then

            // Don't change retcode, may be not handled by extension modules.
            ud_HWCRetcode := pResult^.aData[0]$t_HWCGetHardwareDiagnosisOut.retcode;

            p_UserCalls.p_Callback^.pSvrChCmd.NewInst(pPara,pResult); //Pass on command to extension module

            pResult^.aData[0]$t_HWCGetHardwareDiagnosisOut.retcode := ud_HWCRetcode;

          end_if;
        end_if;

      end_if;

//**********************************************************************************************************************************************************

    CMD_GET_HARDWARE_TREE_ENTRY:

      pResult^.aData$t_HWCGetHardwareTreeEntryOut.retcode := _HWC_RETVAL_ERROR_CLASS_NOT_ONLINE;
      ret_code            := ERROR;

      pStr_HWTRequested   := pPara^.aPara[0]$t_HWCGetHardwareTreeEntryIn.pStr_LastHardewareTreeEntry;

      b_CallThisModule    := TRUE;

      // Check HWT String
      if pStr_HWTRequested & p_ObjectPath then

        // Compare string content
        if _memcmp( ptr1 := pStr_HWTRequested + 2,
                    ptr2 := p_ObjectPath +1,
                    cntr := p_ObjectPath^) = 0 then

          //Check if last call was to Base itself, Compare string length
          if (pStr_HWTRequested$^USINT^ = p_ObjectPath^) then

            //If last call was to base itself, don't call it this time
            b_CallThisModule := FALSE;

            // Last module called was the BusIF Object itself, next module is the 1st behind the extension module
            pPara^.aPara[0]$t_HWCGetHardwareTreeEntryIn.pStr_LastHardewareTreeEntry := NIL;

            if p_UserCalls.p_Callback then
              ret_code := p_UserCalls.p_Callback^.pSvrChCmd.NewInst(pPara,pResult); //Pass on command to extension module

              // if we should quit treating this module special => use standard behavior
              if ret_code = QUIT then
                ret_code := Varan_Base::State.NewInst(pPara,pResult); //Pass on command to base
              end_if;

            else
              pResult^.aData[0]$t_HWCGetHardwareTreeEntryOut.retcode := _HWC_RETVAL_OK_END_OF_LIST;
            end_if;

          elsif (pStr_HWTRequested$^USINT^ > p_ObjectPath^ + 1) then // Must be at least 2 Byte larger, ESCAPE Sequence + Place

            // Check escape sequence
            if ( (pStr_HWTRequested + (p_ObjectPath^) + 2 )^ AND HWT_ESCAPE_SEQU) then // First place after extension module Itself is escape sequence + 1 for addional length byte
              // Last Module must have been a Module behind an extension module

              //If last call was to base itself, don't call it this time
              b_CallThisModule := FALSE;

              // Update index
              pPara^.aPara[0]$t_HWCGetHardwareTreeEntryIn.us_current_index  := p_ObjectPath^ + 3; // Second place after BUSIF Itself is place + 1 for addional length byte
              pPara^.aPara[0]$t_HWCGetHardwareTreeEntryIn.us_current_length := pStr_HWTRequested^ - p_ObjectPath^ - 1;

              //If we have a extension module
              if p_UserCalls.p_Callback then
                ret_code := p_UserCalls.p_Callback^.pSvrChCmd.NewInst(pPara,pResult); //Pass on command to extension module
              else
                ret_code := READY;
                pResult^.aData[0]$t_HWCGetHardwareTreeEntryOut.retcode := _HWC_RETVAL_OK_END_OF_LIST;
              end_if;
            end_if;
          end_if;
        end_if;
      end_if;

      if b_CallThisModule then

        ret_code := Varan_Base::State.NewInst(pPara, pResult);  // Pass on command to base

        // Call conneceted Class for additional info
        if p_UserCalls.p_Callback &
           pResult^.aData[0]$t_HWCGetHardwareTreeEntryOut.pStr_NextHardewareTreeEntry then

          // Update with Requested HWT String with the one returned from Varanbase
          pPara^.aPara[0]$t_HWCGetHardwareTreeEntryIn.pStr_LastHardewareTreeEntry := pResult^.aData[0]$t_HWCGetHardwareTreeEntryOut.pStr_NextHardewareTreeEntry;

          // Don't change retcode, may be not handled by extension modules.
          ud_HWCRetcode := pResult^.aData[0]$t_HWCGetHardwareTreeEntryOut.retcode;

          p_UserCalls.p_Callback^.pSvrChCmd.NewInst(pPara,pResult); //Pass on command to extension module

          pResult^.aData[0]$t_HWCGetHardwareTreeEntryOut.retcode := ud_HWCRetcode;
        end_if;
      end_if;

//**********************************************************************************************************************************************************

   CMD_GET_HW_TIMESTAMP:
      // forward to VM
      ret_code := VaranIn.NewInst(pPara, pResult);

//**********************************************************************************************************************************************************

   CMD_HWC_REQ_PLLNS_REGULATION:
      // forward to VM
      ret_code := VaranIn.NewInst(pPara, pResult);

//**********************************************************************************************************************************************************

  ELSE
    // unknown commands are forwarded to the base
    ret_code := Varan_Base::State.NewInst(pPara, pResult);
  END_CASE;

END_FUNCTION

FUNCTION VIRTUAL GLOBAL BusInterfaceVARAN::GetDeviceID
	VAR_OUTPUT
		output 	: UDINT;
	END_VAR

  output := DeviceIDDiagnosis;

END_FUNCTION

FUNCTION VIRTUAL GLOBAL BusInterfaceVARAN::GetPayloadSupportState
	VAR_OUTPUT
		dRetCode 	: DINT;
	END_VAR

  dRetCode := b_PayloadSupport;

END_FUNCTION

FUNCTION VIRTUAL BusInterfaceVARAN::AddSDORequest
	VAR_INPUT
		pCmdSvr 	: ^SvrChCmd;
		Command 	: HINT;
		Offset 	: UDINT;
		Length 	: UDINT;
		pWriteBuf 	: ^void;
	END_VAR
	VAR_OUTPUT
		sd_retval 	: DINT;
	END_VAR

  // protect via mutex because this can be called from different task priorities
  OS_MT_WAIT(pv_MutexSDOs);

  // if the buffer is full, or the next element in the buffer is already in use
  if (SDOHandling.pWrite^.Command <> 0) then
    sd_retval := -2;
    OS_MT_SIGNAL(pv_MutexSDOs);
    return;
  end_if;

  if pCmdSvr = NIL then
    sd_retval := -3;
    return;
  end_if;

  if Length = 0 then
    sd_retval := -4;
  end_if;

  if Command =_BUS_IF_WRITE_VIA_SDO | Command = _BUS_IF_WRITE_VIA_SDO_CTRL then
    if pWriteBuf = NIL then
      sd_retval := -5;
      return;
    end_if;
  end_if;

  SDOHandling.pWrite^.pCallBackSvr  := pCmdSvr;
  SDOHandling.pWrite^.udLength      := Length;
  SDOHandling.pWrite^.udOffset      := Offset;
  SDOHandling.pWrite^.pWriteData    := pWriteBuf;
  // command is the last thing to store, because it indicates a complete entry
  SDOHandling.pWrite^.Command := Command;

  // we increment our used entries in the buffer (only for debugging)
  SDOHandling.EntriesUsed     += 1;

  // after we successfully added this SDO, set the write pointer to the next element
  if SDOHandling.pWrite = SDOHandling.pLastEntry then
    SDOHandling.pWrite := SDOHandling.pRingBufMemStart;
  else
    SDOHandling.pWrite += sizeof(t_SDORingBufEntry);
  end_if;

  sd_retval := 0;

  OS_MT_SIGNAL(pv_MutexSDOs);

END_FUNCTION

FUNCTION VIRTUAL BusInterfaceVARAN::CyclicSDOHandling
  VAR
		Length 	      : UDINT;
    pRingBufEntry : ^t_SDORingBufEntry;
    pCmdSvr       : ^SvrChCmd;
  	tempCmd       : CmdStruct;
    _result       : results;
    Offset : UDINT;
  END_VAR

  // protect via mutex because this can be called from different task priorities
  OS_MT_WAIT(pv_MutexSDOs);

  //If there is some work todo
  if SDOHandling.EntriesUsed then

    if SDOHandling.pActEntry & SDOHandling.pActEntry^.Command <> 0 then

      pRingBufEntry := SDOHandling.pActEntry;

      //State = 0 ... Start SDO access, 1 ... Get SDO access data and stop SDO
      if SDOHandling.pActEntry^.udState = 0 then

        Length := SDOHandling.pActEntry^.udLength;
        Offset := SDOHandling.pActEntry^.udOffset;

        case SDOHandling.pActEntry^.Command of

          _BUS_IF_READ_VIA_SDO:

            if ChangeAsyRd(Offset:=Offset$UINT,
                           Length:=Length$USINT,
                           RunState:=_BUS_IF_RUN_STATE_CONT_RUN,
                           bIsCtrlACC := FALSE) = FALSE then
              LogError("@009B (BusInterfaceVARAN::CyclicSDOHandling) Error occured at starting the MEM ReadDO");
            end_if;

            SDOHandling.pActEntry^.udState := 1;

          _BUS_IF_READ_VIA_SDO_CTRL:

            if ChangeAsyRd(Offset:=Offset$UINT,
                           Length:=Length$USINT,
                           RunState:=_BUS_IF_RUN_STATE_CONT_RUN,
                           bIsCtrlACC := TRUE) = FALSE then
              LogError("@009B (BusInterfaceVARAN::CyclicSDOHandling) Error occured at starting the CTRL ReadDO");
            end_if;

            SDOHandling.pActEntry^.udState := 1;

          _BUS_IF_WRITE_VIA_SDO:

            _memcpy(ptr1:=AsyMemWriteDO.pData, ptr2:=SDOHandling.pActEntry^.pWriteData, cntr:=SDOHandling.pActEntry^.udLength);

            if ChangeAsyWr(Offset:=Offset$UINT,
                           Length:=Length$USINT,
                           RunState:=_BUS_IF_RUN_STATE_CONT_RUN,
                           bIsCtrlACC := FALSE) = FALSE then
              LogError("@009B (BusInterfaceVARAN::CyclicSDOHandling) Error occured at starting the MEM WriteDO");
            end_if;

            SDOHandling.pActEntry^.udState := 1;

          _BUS_IF_WRITE_VIA_SDO_CTRL:

            _memcpy(ptr1:=AsyCtrlWriteDO.pData, ptr2:=SDOHandling.pActEntry^.pWriteData, cntr:=SDOHandling.pActEntry^.udLength);

            if ChangeAsyWr(Offset:=Offset$UINT,
                           Length:=Length$USINT,
                           RunState:=_BUS_IF_RUN_STATE_CONT_RUN,
                           bIsCtrlACC := TRUE) = FALSE then
              LogError("@009B (BusInterfaceVARAN::CyclicSDOHandling) Error occured at starting the CTRL WriteDO");
            end_if;

            SDOHandling.pActEntry^.udState := 1;

        end_case;

      elsif SDOHandling.pActEntry^.udState = 1 then

        SDOHandling.EntriesUsed -= 1;

        // Call the corresponding function in the operator class
        tempCmd.uiCmd := _BUS_IF_SDO_RESPONSE;
        tempCmd.aPara[0] := SDOHandling.pActEntry^.Command$DINT;
        tempCmd.aPara[1] := SDOHandling.pActEntry^.udOffset$DINT;
        tempCmd.aPara[2] := SDOHandling.pActEntry^.udLength$DINT;

        tempCmd.aPara[3] := 0;

        case SDOHandling.pActEntry^.Command of

          _BUS_IF_READ_VIA_SDO:

            tempCmd.aPara[4] := AsyMemReadDO.pData$DINT;
            tempCmd.aPara[5] := AsyMemReadDO.Length;

          _BUS_IF_READ_VIA_SDO_CTRL:

            tempCmd.aPara[4] := AsyCtrlReadDO.pData$DINT;
            tempCmd.aPara[5] := AsyCtrlReadDO.Length;

          _BUS_IF_WRITE_VIA_SDO:

            tempCmd.aPara[4] := NIL$DINT;
            tempCmd.aPara[5] := 0;

          _BUS_IF_WRITE_VIA_SDO_CTRL:

            tempCmd.aPara[4] := NIL$DINT;
            tempCmd.aPara[5] := 0;

        end_case;

        pCmdSvr := pRingBufEntry^.pCallBackSvr;

        if pCmdSvr$pVirtualBase^.NewInst(#tempCmd, #_result) <> READY then
          LogError("@0099 (BusInterfaceVARAN::CyclicSDOHandling) SDO Error: Error of module at place 0x{0} while receiving the SDO reponse (which was an ErrorCode)");
        end_if;

        // the entry in the ringbuffer is free
        pRingBufEntry^.Command := 0;

        //Stop the DOs
        if ChangeAsyRd(Offset:=0,
                       Length:=0,
                       RunState:=_BUS_IF_RUN_STATE_NO_RUN,
                       bIsCtrlACC := TRUE) = FALSE then
          LogError("@0769 (BusInterfaceVARAN::CyclicSDOHandling) Error occured at starting the CTRL ReadDO");
        end_if;

        if ChangeAsyRd(Offset:=0,
                       Length:=0,
                       RunState:=_BUS_IF_RUN_STATE_NO_RUN,
                       bIsCtrlACC := FALSE) = FALSE then
          LogError("@076A (BusInterfaceVARAN::CyclicSDOHandling) Error occured at starting the MEM ReadDO");
        end_if;

        if ChangeAsyWr(Offset:=0,
                       Length:=0,
                       RunState:=_BUS_IF_RUN_STATE_NO_RUN,
                       bIsCtrlACC := TRUE) = FALSE then
          LogError("@076B (BusInterfaceVARAN::CyclicSDOHandling) Error occured at starting the CTRL WriteDO");
        end_if;

        if ChangeAsyWr(Offset:=0,
                       Length:=0,
                       RunState:=_BUS_IF_RUN_STATE_NO_RUN,
                       bIsCtrlACC := FALSE) = FALSE then
          LogError("@076D (BusInterfaceVARAN::CyclicSDOHandling) Error occured at starting the MEM WriteDO");
        end_if;

        SDOHandling.pActEntry^.udState := 0;

        // after we successfully added this SDO, set the read pointer to the next element
        if SDOHandling.pActEntry = SDOHandling.pLastEntry then
          SDOHandling.pActEntry := SDOHandling.pRingBufMemStart;
        else
          SDOHandling.pActEntry += sizeof(t_SDORingBufEntry);
        end_if;

      end_if;
    end_if;
  end_if;

  OS_MT_SIGNAL(pv_MutexSDOs);

END_FUNCTION

FUNCTION VIRTUAL BusInterfaceVARAN::ChangeAsyRd
	VAR_INPUT
		Offset 	: HINT;
		Length 	: USINT;
		RunState 	: t_BusIFRunState;
		bIsCtrlACC 	: BOOL;
	END_VAR
	VAR_OUTPUT
		Success 	: BOOL;
	END_VAR
  VAR
    dataUPDATEDO    : t_UpdateDOCfg;
  	tempCmd         : CmdStruct;
    _result         : results;
    dataSETRUNSTATE : t_SetRunStateCfg;
  END_VAR

  // if length = zero we may just want to stop the DO
  if Length then

    if bIsCtrlACC then
      AsyCtrlReadDO.Offset := Offset;
      AsyCtrlReadDO.Length := Length;

      dataUPDATEDO.Handle               := AsyCtrlReadDO.Handle;
      dataUPDATEDO.ud_addressoff_read   := AsyCtrlReadDO.Offset;
      dataUPDATEDO.ud_length_read       := AsyCtrlReadDO.Length;

    else
      AsyMemReadDO.Offset := Offset;
      AsyMemReadDO.Length := Length;

      dataUPDATEDO.Handle               := AsyMemReadDO.Handle;
      dataUPDATEDO.ud_addressoff_read   := AsyMemReadDO.Offset;
      dataUPDATEDO.ud_length_read       := AsyMemReadDO.Length;
    end_if;

    tempCmd.uiCmd         := _BUS_IF_UPDATE_DO;
    tempCmd.aPara[0]      := (#dataUPDATEDO)$DINT;

    CallCommand.NewInst(pPara:=#tempCmd, pResult:=#_result);
    if _result.aData[0]$t_BusIFRetvalErrorcode <> _BUS_IF_RETVAL_OK then
      LogError("@007C (BusInterfaceVARAN::ChangeAsyRd) Failed to change asynchron read access");
    end_if;
  end_if;

  // set runstate
  if bIsCtrlACC then
    dataSETRUNSTATE.Handle      := AsyCtrlReadDO.Handle;
  else
    dataSETRUNSTATE.Handle      := AsyMemReadDO.Handle;
  end_if;

  dataSETRUNSTATE.NewRunState := RunState;

  tempCmd.uiCmd         := _BUS_IF_SET_RUN_STATE;
  tempCmd.aPara[0]      := (#dataSETRUNSTATE)$DINT;

  CallCommand.NewInst(pPara:=#tempCmd, pResult:=#_result);

  if _result.aData[0]$t_BusIFRetvalErrorcode <> _BUS_IF_RETVAL_OK then
    LogError("@007D (BusInterfaceVARAN::ChangeAsyRd) Error changing the run state of the asynchron read access!");
  end_if;

  Success := TRUE;

END_FUNCTION

FUNCTION VIRTUAL BusInterfaceVARAN::ChangeAsyWr
	VAR_INPUT
		Offset 	: HINT;
		Length 	: USINT;
		RunState 	: t_BusIFRunState;
		bIsCtrlACC 	: BOOL;
	END_VAR
	VAR_OUTPUT
		Success 	: BOOL;
	END_VAR
  VAR
    dataUPDATEDO    : t_UpdateDOCfg;
  	tempCmd         : CmdStruct;
    _result         : results;
    dataSETRUNSTATE : t_SetRunStateCfg;
  END_VAR

  // if length = zero we may just want to stop the DO
  if Length then

    if bIsCtrlACC then
      AsyCtrlWriteDO.Offset := Offset;
      AsyCtrlWriteDO.Length := Length;

      dataUPDATEDO.Handle               := AsyCtrlWriteDO.Handle;
      dataUPDATEDO.ud_addressoff_write  := AsyCtrlWriteDO.Offset;
      dataUPDATEDO.ud_length_write      := AsyCtrlWriteDO.Length;

    else
      AsyMemWriteDO.Offset := Offset;
      AsyMemWriteDO.Length := Length;

      dataUPDATEDO.Handle               := AsyMemWriteDO.Handle;
      dataUPDATEDO.ud_addressoff_write  := AsyMemWriteDO.Offset;
      dataUPDATEDO.ud_length_write      := AsyMemWriteDO.Length;

    end_if;

    tempCmd.uiCmd         := _BUS_IF_UPDATE_DO;
    tempCmd.aPara[0]      := (#dataUPDATEDO)$DINT;

    CallCommand.NewInst(pPara:=#tempCmd, pResult:=#_result);
    if _result.aData[0]$t_BusIFRetvalErrorcode <> _BUS_IF_RETVAL_OK then
      LogError("@007F (BusInterfaceVARAN::ChangeAsyWr) Failed to change asynchron write access");
    end_if;
  end_if;

  // set runstate
  if bIsCtrlACC then
    dataSETRUNSTATE.Handle      := AsyCtrlWriteDO.Handle;
  else
    dataSETRUNSTATE.Handle      := AsyMemWriteDO.Handle;
  end_if;

  dataSETRUNSTATE.NewRunState := RunState;

  tempCmd.uiCmd         := _BUS_IF_SET_RUN_STATE;
  tempCmd.aPara[0]      := (#dataSETRUNSTATE)$DINT;

  CallCommand.NewInst(pPara:=#tempCmd, pResult:=#_result);

  if _result.aData[0]$t_BusIFRetvalErrorcode <> _BUS_IF_RETVAL_OK then
    LogError("@0080 (BusInterfaceVARAN::ChangeAsyWr) Error changing the run state of the asynchron write access!");
  end_if;

  Success := TRUE;

END_FUNCTION

FUNCTION VIRTUAL BusInterfaceVARAN::SendPostInitFinished
	VAR_INPUT
		DisableThisObject 	: BOOL;(* := FALSE *)
	END_VAR
  VAR
  	tempCmd         : CmdStruct;
    _result         : results;
  END_VAR

  b_PostInitFinished := TRUE;
  tempCmd.uiCmd := _BUS_IF_POST_INIT_FINISHED;
  CallCommand.NewInst(pPara:=#tempCmd, pResult:=#_result);

  if _result.aData[0]$t_BusIFRetvalErrorcode <> _BUS_IF_RETVAL_OK then
    LogError("@00D8 (BusInterfaceVARAN::SendPostInitFinished) Failed to set the post init to finished via bus interface!");
  end_if;

  if DisableThisObject then
    // tell the manager that we don't need to be called for rt syncing
    tempCmd.uiCmd := _BUS_IF_RT_SYNC_READY;
    CallCommand.NewInst(pPara:=#tempCmd, pResult:=#_result);

    if _result.aData[0]$t_BusIFRetvalErrorcode <> _BUS_IF_RETVAL_OK then
      LogError("@00D9 (BusInterfaceVARAN::CyWork) Failed to set rt sync ready via bus interface!");
    end_if;
  end_if;

END_FUNCTION

FUNCTION VIRTUAL BusInterfaceVARAN::SimulateSDIASManagerCywork
VAR
	tempCmd           : CmdStruct;
  _result           : results;
  RetcodeIPR        : iprStates;
END_VAR

  case eSdiasManagerInitSSW of
//**********************************************************************************************************************************************************
    t_SdiasManagerInitSSW::_StartInit:

      // remember when we started (for timeout and init time measure)
      InitStartTime := ops.tAbsolute;

      // check if we have a user class
      if p_UserCalls.p_Callback = NIL then
        // we already have a log entry from the constructor
        State := _CallBackError;
        LogError("@076E (BusInterfaceVARAN::SimulateSDIASManagerCywork) Pointer to user callback is invalid");
        eErrorInitStep := eSdiasManagerInitSSW;
        eSdiasManagerInitSSW := _PrepareError;
        return;
      end_if;

      //Go on with initialisation
      eSdiasManagerInitSSW := _InitAccesses;

//**********************************************************************************************************************************************************
    t_SdiasManagerInitSSW::_InitAccesses:

      // call operator, who returns the init state (busy = call me again, error = error occured/cancel init, ready = init successfully finished)
      if p_UserCalls.p_Callback then
        // Call the corresponding function in the operator class
        tempCmd.uiCmd := _BUS_IF_INIT_ACCESSES;
        RetcodeIPR := p_UserCalls.p_Callback^.pSvrChCmd.NewInst(#tempCmd,#_result);
      else
        RetcodeIPR := READY;
      end_if;

      if RetcodeIPR = READY then
        eSdiasManagerInitSSW := t_SdiasManagerInitSSW::_FinishInitialisation;
      elsif RetcodeIPR = ERROR then
        eErrorInitStep := eSdiasManagerInitSSW;
        eSdiasManagerInitSSW := t_SdiasManagerInitSSW::_PrepareError;
      end_if;

//**********************************************************************************************************************************************************
    t_SdiasManagerInitSSW::_FinishInitialisation:

      // tell the manager that we're finished with initializing, otherwise realtime will not be called
      if b_PostInitFinished = FALSE then
        SendPostInitFinished();
      end_if;

      //Enable the DOs in realtime
      eSdiasManagerInitSSW := _CallHwConnect;

//**********************************************************************************************************************************************************
    t_SdiasManagerInitSSW::_CallHwConnect:

      //Do nothing here, work is done in realtime (so that DOs will be started in the correct task

//**********************************************************************************************************************************************************
    t_SdiasManagerInitSSW::_ModuleInitialisation:

      // call operator, who returns the init state (busy = call me again, error = error occured/cancel init, ready = init successfully finished)
      if p_UserCalls.p_Callback then
        // Call the corresponding function in the operator class
        tempCmd.uiCmd := _BUS_IF_INIT_MODULE;
        RetcodeIPR := p_UserCalls.p_Callback^.pSvrChCmd.NewInst(#tempCmd,#_result);
      else
        RetcodeIPR := READY;
      end_if;

      if RetcodeIPR = READY then
        eSdiasManagerInitSSW := t_SdiasManagerInitSSW::_InitFinished;

        if bSendRtSyncReady = FALSE then

          bSendRtSyncReady := TRUE;
          //Finish init
          tempCmd.uiCmd := _BUS_IF_RT_SYNC_READY;
          CallCommand.NewInst(pPara:=#tempCmd, pResult:=#_result);

          if _result.aData[0]$t_BusIFRetvalErrorcode <> _BUS_IF_RETVAL_OK then
            LogError("@00D9 (BusInterfaceVARAN::CyWork) Failed to set rt sync ready via bus interface!");
          end_if;
        end_if;

      elsif RetcodeIPR = ERROR then
        eErrorInitStep := eSdiasManagerInitSSW;
        eSdiasManagerInitSSW := t_SdiasManagerInitSSW::_PrepareError;
      end_if;

//**********************************************************************************************************************************************************
    t_SdiasManagerInitSSW::_InitFinished:

      p_UserCalls.p_UpdateCy^.CyWork(EAX:=0);

//**********************************************************************************************************************************************************
    t_SdiasManagerInitSSW::_PrepareError:

    // tell the manager that we're finished with initializing
    if b_PostInitFinished = FALSE then
      SendPostInitFinished(DisableThisObject:=TRUE);
    end_if;

    //Sets a required error if the module is required
    SetRequiredError();

    eSdiasManagerInitSSW := _ErrorOccured;

//**********************************************************************************************************************************************************
    t_SdiasManagerInitSSW::_ErrorOccured:
      // do nothing here
      return;

  end_case;

  //Always call SDO Handling
  CyclicSDOHandling();

END_FUNCTION

FUNCTION VIRTUAL BusInterfaceVARAN::SetRequiredError
  VAR
  	tempCmd         : CmdStruct;
    _result         : results;
  END_VAR

  if Required then

    // set required error
    tempCmd.uiCmd     := _BUS_IF_SET_REQUIRED_ERROR;

    CallCommand.NewInst(pPara:=#tempCmd, pResult:=#_result);
    if _result.aData[0]$t_BusIFRetvalErrorcode <> _BUS_IF_RETVAL_OK then
      LogError("@00A1 (BusInterfaceVARAN::SetRequiredError) Failed to set required error");
    end_if;
  end_if;

END_FUNCTION

FUNCTION VIRTUAL BusInterfaceVARAN::SimulateSDIASManagerRtwork
VAR
	tempCmd     : CmdStruct;
  _result     : results;
END_VAR

  case eSdiasManagerRTSSW of
  	t_SdiasManagerRtSSW::_RtIdle: // nothing
  	t_SdiasManagerRtSSW::_CreateAndModifyDOs: //nothing to do here
  	t_SdiasManagerRtSSW::_Wait4DOs:
  	t_SdiasManagerRtSSW::_Wait4PllSync:
  	t_SdiasManagerRtSSW::_Wait2Ticks:
  	t_SdiasManagerRtSSW::_CntDownSyncStart:
  	t_SdiasManagerRtSSW::_PreOperationalWait4DataReady:
  	t_SdiasManagerRtSSW::_PreOperational:
  	t_SdiasManagerRtSSW::_Operational:
  end_case;

  if eSdiasManagerInitSSW = _CallHwConnect then

    if bCallHwConnectInRT then
      bCallHwConnectInRT := FALSE;

      // Call the corresponding function in the operator class
      tempCmd.uiCmd := _BUS_IF_HWCONNECT;
      p_UserCalls.p_Callback^.pSvrChCmd.NewInst(#tempCmd,#_result);

      eSdiasManagerInitSSW := _ModuleInitialisation;

      if _result.aData[0] then
        return;
      end_if;
    end_if;
  end_if;

END_FUNCTION
